Fanuc KAREL source: KT00756.KL

PROGRAM KT00756
%NOLOCKGROUP
VAR
  B1: BOOLEAN
  B2: BOOLEAN
  OUT: INTEGER
BEGIN
  B1 = TRUE
  B2 = FALSE
  B1 = TRUE
  B2 = FALSE
  OUT = ABS(B1)
END KT00756
